// TIA Portal V21 export
// export: Created 2026-11-08T21:21:37.5603302Z, ExportSetting WithDefaults, DisplayName Totally Integrated Automation Portal, DisplayVersion V21 Update 3, DisplayName STEP 7 Professional, DisplayVersion V21 Update 3, DisplayName STEP 7 Safety, DisplayVersion V21, DisplayName Tech WebApplication, DisplayVersion V21, DisplayName WinCC Basic/Comfort/Advanced, DisplayVersion V21 Update 3, DisplayName WinCC Unified, DisplayVersion V21 Update 3
DATA_BLOCK "DB_StlInner"   // DB7
VERSION : 0.1
// stored: AutoNumber true, DBAccessibleFromOPCUA true, DBAccessibleFromWebserver true, InstanceOfName FB_StlInner, InstanceOfType FB
"FB_StlInner"
   // VAR_INPUT
   //    start : Bool;
   // END_VAR
   // VAR_OUTPUT
   //    cnt : Int;
   // END_VAR
   // VAR
   //    n : Int;
   // END_VAR
BEGIN
END_DATA_BLOCK
